// TwinCAT 3 PLC project Untitled1
// ProgramVersion: 3.1.4024.0
// libraries:
//   Tc2_Math, * (Beckhoff Automation GmbH)
//   Tc2_Standard, * (Beckhoff Automation GmbH)
//   Tc2_System, * (Beckhoff Automation GmbH)
//   Tc3_Module, * (Beckhoff Automation GmbH)
//   Tc2_MC2, * (Beckhoff Automation GmbH)
//   Tc2_MC2_Camming, * (Beckhoff Automation GmbH)
// project tree:
//   DUTs/ E_CamApplicationError.TcDUT, E_CamErrorSource.TcDUT, E_CamMachineState.TcDUT, E_CamProcessPhase.TcDUT, ST_CamCommands.TcDUT, ST_CamDerivedGeometry.TcDUT, ST_CamRecipe.TcDUT, ST_CamScope.TcDUT, ST_CamStatus.TcDUT
//   GVLs/ GVL_CamControl.TcGVL, GVL_Motion.TcGVL
//   / PlcTask.TcTTO (not stored)
//   POUs/Cam/ FB_CamMachine.TcPOU, FB_CamProfileBuilder.TcPOU, FB_CamRecipeValidator.TcPOU, FB_ElectronicCam.TcPOU, F_MakeCamPoint.TcPOU
//   POUs/Axis_test/ Axis_test.TcPOU, FB_AxisPositionTest.TcPOU
//   POUs/ MAIN.TcPOU
// real-time tasks:
//   TASK PlcTask: cycle T#10ms, priority 20, ADS port 350
// motion (NC):
//   TASK NC-Task 1 SAF: cycle T#2ms, priority 4, ADS port 501
//   TASK NC-Task 1 SVB: cycle T#10ms, priority 8, ADS port 511
//   AXIS Axis 1 (id 1)
//     OtherSettings: AllowMotionCmdToSlave=true
//     encoder EncType=19
//       EncPara: MaxCount=#xffffffff
//     drive DrvType=16
//       DrvPara: MaxCount=#xffffffff
//         Analog: TorqueSetpointScale=10, ScaleFactorActTorque=0.1
//         TimeComp: TaskDelayCycles=1
//     controller CtrType=1
//       CtrPara: PriorControlFactor=1
//         Observer: BandWidth=20
//   AXIS Axis 2 (id 2)
//     OtherSettings: AllowMotionCmdToSlave=true
//     encoder EncType=19
//       EncPara: MaxCount=#xffffffff
//     drive DrvType=16
//       DrvPara: MaxCount=#xffffffff
//         Analog: TorqueSetpointScale=10, ScaleFactorActTorque=0.1
//         TimeComp: TaskDelayCycles=1
//     controller CtrType=1
//       CtrPara: PriorControlFactor=1
//         Observer: BandWidth=20
// I/O:
//   DEVICE Device 3 (EtherCAT), AmsNetId 5.57.253.57.4.1
//     Drive 1 (INVT_DA180_114) [DA180-N EtherCAT(CoE) Drive]
//     Drive 2 (INVT_DA200A_EtherCAT_101) [INVT_DA200A_EtherCAT_1.0.1.0]
//     Term 3 (EK1100) [EK1100 EtherCAT Coupler (2A E-Bus)]
//       Term 4 (EL3164) [EL3164 4Ch. Ana. Input 0-10V]
//       Term 5 (EL9011) [EL9011 End Terminal]
// variable links:
//   NC-Task 1 SAF/Axes/Axis 1 <-> Device 3 (EtherCAT)/Drive 1 (INVT_DA180_114)
//     Drive/Inputs/In/nDataIn3[0] <-> DI Inputs/Torque Actual Value
//     Drive/Inputs/In/nDcOutputTime <-> InfoData/DcOutputShift
//     Drive/Inputs/In/nState1 <-> DI Inputs/Status Word
//     Drive/Inputs/In/nState2 <-> DI Inputs/Status Word @bit 8
//     Drive/Inputs/In/nState4 @bit 1 <-> WcState/InputToggle
//     Drive/Inputs/In/nState4 <-> WcState/WcState
//     Drive/Inputs/In/nState5 <-> DI Inputs/Operation Mode Display
//     Drive/Outputs/Out/nCtrl1 <-> DO Outputs/Control Word
//     Drive/Outputs/Out/nCtrl2 <-> DO Outputs/Control Word @bit 8
//     Drive/Outputs/Out/nCtrl5 <-> DO Outputs/Mode of Operation
//     Drive/Outputs/Out/nDataOut1 <-> DO Outputs/Target Position
//     Drive/Outputs/Out/nDataOut2 <-> DO Outputs/Target Velocity
//     Drive/Outputs/Out/nDataOut4[0] <-> DO Outputs/Target torque
//     Enc/Inputs/In/nDataIn1 <-> DI Inputs/Position Actual Value
//     Enc/Inputs/In/nDataIn3 <-> DI Inputs/Touch Probe Value
//     Enc/Inputs/In/nDataIn7 <-> DI Inputs/Speed Actual Value
//     Enc/Inputs/In/nDcInputTime <-> InfoData/DcInputShift
//     Enc/Inputs/In/nState4 @bit 1 <-> WcState/InputToggle
//     Enc/Inputs/In/nState4 <-> WcState/WcState
//     Enc/Inputs/In/nState5 <-> DI Inputs/Touch Probe Status
//     Enc/Inputs/In/nState6 <-> DI Inputs/Touch Probe Status @bit 8
//     Enc/Outputs/Out/nCtrl5 <-> DO Outputs/Touch probe control
//     Enc/Outputs/Out/nCtrl6 <-> DO Outputs/Touch probe control @bit 8
//   NC-Task 1 SAF/Axes/Axis 2 <-> Device 3 (EtherCAT)/Drive 2 (INVT_DA200A_EtherCAT_101)
//     Drive/Inputs/In/nDataIn3[0] <-> Inputs/Torque Actual Value
//     Drive/Inputs/In/nDcOutputTime <-> InfoData/DcOutputShift
//     Drive/Inputs/In/nState1 <-> Inputs/Status Word
//     Drive/Inputs/In/nState2 <-> Inputs/Status Word @bit 8
//     Drive/Inputs/In/nState4 @bit 1 <-> WcState/InputToggle
//     Drive/Inputs/In/nState4 <-> WcState/WcState
//     Drive/Inputs/In/nState5 <-> Inputs/Operation Mode Display
//     Drive/Outputs/Out/nCtrl1 <-> Outputs/Control Word
//     Drive/Outputs/Out/nCtrl2 <-> Outputs/Control Word @bit 8
//     Drive/Outputs/Out/nCtrl5 <-> Outputs/Mode of Operation
//     Drive/Outputs/Out/nDataOut1 <-> Outputs/Target Position
//     Drive/Outputs/Out/nDataOut2 <-> Outputs/Target Velocity
//     Drive/Outputs/Out/nDataOut4[0] <-> Outputs/Target torque
//     Enc/Inputs/In/nDataIn1 <-> Inputs/Position Actual Value
//     Enc/Inputs/In/nDataIn3 <-> Inputs/Touch Probe 1 Positive value
//     Enc/Inputs/In/nDataIn7 <-> Inputs/Velocity Actual Value
//     Enc/Inputs/In/nDcInputTime <-> InfoData/DcInputShift
//     Enc/Inputs/In/nState4 @bit 1 <-> WcState/InputToggle
//     Enc/Inputs/In/nState4 <-> WcState/WcState
//     Enc/Inputs/In/nState5 <-> Inputs/Touch Probe Status
//     Enc/Inputs/In/nState6 <-> Inputs/Touch Probe Status @bit 8
//     Enc/Outputs/Out/nCtrl5 <-> Outputs/Touch probe control
//     Enc/Outputs/Out/nCtrl6 <-> Outputs/Touch probe control @bit 8
//   Untitled1/Untitled1 Instance <-> NC-Task 1 SAF/Axes/Axis 1
//     PlcTask Inputs/GVL_Motion.gAxisConveyor.NcToPlc <-> Outputs/ToPlc
//     PlcTask Outputs/GVL_Motion.gAxisConveyor.PlcToNc <-> Inputs/FromPlc
//   Untitled1/Untitled1 Instance <-> NC-Task 1 SAF/Axes/Axis 2
//     PlcTask Inputs/GVL_Motion.gAxisCutter.NcToPlc <-> Outputs/ToPlc
//     PlcTask Outputs/GVL_Motion.gAxisCutter.PlcToNc <-> Inputs/FromPlc

// ---- DUTs/E_CamApplicationError.TcDUT
TYPE E_CamApplicationError :
(
    CAM_ERROR_NONE := 0,
    CAM_ERROR_COMMAND_NOT_ALLOWED,
    CAM_ERROR_NOT_REFERENCED,
    CAM_ERROR_RECIPE_PITCH,
    CAM_ERROR_RECIPE_CONVEYOR_VELOCITY,
    CAM_ERROR_RECIPE_CUT_VELOCITY,
    CAM_ERROR_RECIPE_EDGE_LENGTH,
    CAM_ERROR_RECIPE_PHASE_ORDER,
    CAM_ERROR_RECIPE_SYNC_SPACE,
    CAM_ERROR_RECIPE_RETURN_SPACE,
    CAM_ERROR_RECIPE_DYNAMICS,
    CAM_ERROR_AXIS_POWER,
    CAM_ERROR_AXIS_REFERENCE,
    CAM_ERROR_CAM_BUILD,
    CAM_ERROR_CAM_LOAD,
    CAM_ERROR_CAM_CHARACTERISTICS,
    CAM_ERROR_CAM_IN,
    CAM_ERROR_MASTER_MOVE,
    CAM_ERROR_MASTER_STOP,
    CAM_ERROR_CAM_OUT,
    CAM_ERROR_SLAVE_RETURN,
    CAM_ERROR_AXIS_RESET
);
END_TYPE

// ---- DUTs/E_CamErrorSource.TcDUT
TYPE E_CamErrorSource :
(
    CAM_SOURCE_NONE := 0,
    CAM_SOURCE_RECIPE,
    CAM_SOURCE_MASTER_AXIS,
    CAM_SOURCE_SLAVE_AXIS,
    CAM_SOURCE_TABLE_LOAD,
    CAM_SOURCE_TABLE_CHARACTERISTICS,
    CAM_SOURCE_CAM_IN,
    CAM_SOURCE_CAM_OUT
);
END_TYPE

// ---- DUTs/E_CamMachineState.TcDUT
TYPE E_CamMachineState :
(
    CAM_STATE_DISABLED := 0,
    CAM_STATE_POWERING,
    CAM_STATE_IDLE,
    CAM_STATE_REFERENCING_MASTER,
    CAM_STATE_REFERENCING_SLAVE,
    CAM_STATE_BUILDING_TABLE,
    CAM_STATE_LOADING_TABLE,
    CAM_STATE_READY,
    CAM_STATE_CAMMING_IN,
    CAM_STATE_STARTING_MASTER,
    CAM_STATE_RUNNING,
    CAM_STATE_STOPPING_MASTER,
    CAM_STATE_RELEASING_STOP,
    CAM_STATE_CAMMING_OUT,
    CAM_STATE_RETURNING_SLAVE,
    CAM_STATE_RESETTING,
    CAM_STATE_FAULT
);
END_TYPE

// ---- DUTs/E_CamProcessPhase.TcDUT
TYPE E_CamProcessPhase :
(
    CAM_PHASE_DISABLED := 0,
    CAM_PHASE_PREPARE,
    CAM_PHASE_APPROACH,
    CAM_PHASE_FIRST_EDGE,
    CAM_PHASE_EXIT_FIRST_EDGE,
    CAM_PHASE_SYNCHRONOUS,
    CAM_PHASE_ENTER_SECOND_EDGE,
    CAM_PHASE_SECOND_EDGE,
    CAM_PHASE_RETURN,
    CAM_PHASE_DWELL
);
END_TYPE

// ---- DUTs/ST_CamCommands.TcDUT
TYPE ST_CamCommands :
STRUCT
    bEnable : BOOL;
    bReference : BOOL;
    bApplyRecipe : BOOL;
    bStart : BOOL;
    bStop : BOOL;
    bReset : BOOL;
END_STRUCT
END_TYPE

// ---- DUTs/ST_CamDerivedGeometry.TcDUT
TYPE ST_CamDerivedGeometry :
STRUCT
    lrCutMasterDistance : LREAL;
    lrFirstSlope : LREAL;
    lrSecondSlope : LREAL;
    lrFirstEdgeEnd : LREAL;
    lrExitBlendEnd : LREAL;
    lrEntryBlendStart : LREAL;
    lrSecondEdgeEnd : LREAL;
    lrClearanceRelative : LREAL;
    lrFirstStartY : LREAL;
    lrFirstEndY : LREAL;
    lrExitEndY : LREAL;
    lrEntryStartY : LREAL;
    lrSecondStartY : LREAL;
    lrSecondEndY : LREAL;
    lrMasterStopDistance : LREAL;
    lrStopWindowMargin : LREAL;
END_STRUCT
END_TYPE

// ---- DUTs/ST_CamRecipe.TcDUT
TYPE ST_CamRecipe :
STRUCT
    lrObjectPitch : LREAL := 500.0;
    lrConveyorVelocity : LREAL := 100.0;
    lrCutVelocity : LREAL := 50.0;
    lrObjectEdgeLength : LREAL := 25.0;
    lrFirstEdgeStart : LREAL := 100.0;
    lrSecondEdgeStart : LREAL := 300.0;
    lrBlendMasterDistance : LREAL := 20.0;
    lrReturnEndPhase : LREAL := 480.0;
    lrMasterAcceleration : LREAL := 500.0;
    lrMasterDeceleration : LREAL := 500.0;
    lrMasterJerk : LREAL := 5000.0;
    lrMaxSlaveVelocity : LREAL := 600.0;
    lrMaxSlaveAcceleration : LREAL := 1600.0;
    lrMaxSlaveJerk : LREAL := 12000.0;
    lrRecoveryVelocity : LREAL := 100.0;
    lrRecoveryAcceleration : LREAL := 500.0;
    lrRecoveryDeceleration : LREAL := 500.0;
    lrRecoveryJerk : LREAL := 5000.0;
    lrPositionTolerance : LREAL := 0.1;
END_STRUCT
END_TYPE

// ---- DUTs/ST_CamScope.TcDUT
TYPE ST_CamScope :
STRUCT
    lrMasterSetPosition : LREAL;
    lrMasterActualPosition : LREAL;
    lrMasterSetVelocity : LREAL;
    lrMasterActualVelocity : LREAL;
    lrMasterPhase : LREAL;
    lrSlaveSetPosition : LREAL;
    lrSlaveActualPosition : LREAL;
    lrSlaveSetVelocity : LREAL;
    lrSlaveActualVelocity : LREAL;
    lrExpectedSlaveVelocity : LREAL;
    lrObjectRelativePosition : LREAL;
    eMachineState : E_CamMachineState;
    eProcessPhase : E_CamProcessPhase;
    bCamActive : BOOL;
    bRecipeLoaded : BOOL;
    eApplicationError : E_CamApplicationError;
    udiMotionErrorID : UDINT;
END_STRUCT
END_TYPE

// ---- DUTs/ST_CamStatus.TcDUT
TYPE ST_CamStatus :
STRUCT
    eState : E_CamMachineState;
    eProcessPhase : E_CamProcessPhase;
    bPowerEnabled : BOOL;
    bReferenced : BOOL;
    bRecipeLoaded : BOOL;
    bCamActive : BOOL;
    bRunning : BOOL;
    bBusy : BOOL;
    eApplicationError : E_CamApplicationError;
    eErrorSource : E_CamErrorSource;
    udiMotionErrorID : UDINT;
    lrCalculatedMaxSlaveVelocity : LREAL;
    lrCalculatedMaxSlaveAcceleration : LREAL;
    lrCalculatedMaxSlaveJerk : LREAL;
    lrCalculatedFaultStopSlaveAcceleration : LREAL;
    lrCalculatedFaultStopSlaveJerk : LREAL;
END_STRUCT
END_TYPE

// ---- GVLs/GVL_CamControl.TcGVL
{attribute 'qualified_only'}
VAR_GLOBAL
    stCommands : ST_CamCommands;
    stRecipe : ST_CamRecipe;
    stStatus : ST_CamStatus;
    stScope : ST_CamScope;
END_VAR

// ---- GVLs/GVL_Motion.TcGVL
{attribute 'qualified_only'}
VAR_GLOBAL
    gAxisConveyor : AXIS_REF;
    gAxisCutter : AXIS_REF;
END_VAR

// ---- POUs/Cam/FB_CamMachine.TcPOU
FUNCTION_BLOCK FB_CamMachine
VAR_INPUT
    stCommands : ST_CamCommands;
    stRecipe : ST_CamRecipe;
END_VAR
VAR_IN_OUT
    AxisConveyor : AXIS_REF;
    AxisCutter : AXIS_REF;
END_VAR
VAR_OUTPUT
    stStatus : ST_CamStatus;
    stScope : ST_CamScope;
END_VAR
VAR CONSTANT
    c_nCamTableIdA : MC_CAM_ID := 1;
    c_nCamTableIdB : MC_CAM_ID := 2;
    // Commissioned application limits; NC/drive limits must be no lower.
    c_lrMachineMaxSlaveVelocity : LREAL := 600.0;
    c_lrMachineMaxSlaveAcceleration : LREAL := 1600.0;
    c_lrMachineMaxSlaveJerk : LREAL := 12000.0;
    // Conservative controlled stop used only after a runtime fault.
    c_lrFaultStopDeceleration : LREAL := 15.0;
    c_lrFaultStopJerk : LREAL := 50.0;
END_VAR
VAR
    eState : E_CamMachineState := CAM_STATE_DISABLED;
    eProcessPhase : E_CamProcessPhase := CAM_PHASE_DISABLED;

    rtReference : R_TRIG;
    rtApplyRecipe : R_TRIG;
    rtStart : R_TRIG;
    rtStop : R_TRIG;
    rtReset : R_TRIG;

    fbPowerConveyor : MC_Power;
    fbPowerCutter : MC_Power;
    fbSetPositionConveyor : MC_SetPosition;
    fbSetPositionCutter : MC_SetPosition;
    fbResetConveyor : MC_Reset;
    fbResetCutter : MC_Reset;
    fbMoveConveyor : MC_MoveVelocity;
    fbStopConveyor : MC_Stop;
    fbReturnCutter : MC_MoveAbsolute;

    fbRecipeValidator : FB_CamRecipeValidator;
    fbProfileBuilder : FB_CamProfileBuilder;
    fbElectronicCam : FB_ElectronicCam;

    stPowerOptions : ST_PowerOptions;
    stSetPositionConveyorOptions : ST_SetPositionOptions;
    stSetPositionCutterOptions : ST_SetPositionOptions;
    stMoveConveyorOptions : ST_MoveOptions;
    stStopConveyorOptions : ST_MoveOptions;
    stReturnCutterOptions : ST_MoveOptions;

    stPendingRecipe : ST_CamRecipe;
    stActiveRecipe : ST_CamRecipe;
    stDerived : ST_CamDerivedGeometry;
    stCamRef : MC_CAM_REF;

    bPowerRequest : BOOL;
    bReferenced : BOOL;
    bRecipeLoaded : BOOL;
    bStopRequested : BOOL;
    bResetInProgress : BOOL;
    bFaultStop : BOOL;
    bForcePowerOff : BOOL;
    usiBuildState : USINT;

    nActiveCamTableId : MC_CAM_ID := 1;
    nCandidateCamTableId : MC_CAM_ID := 2;
    nCamCommandTableId : MC_CAM_ID := 1;

    bSetPositionConveyorExecute : BOOL;
    bSetPositionCutterExecute : BOOL;
    bResetConveyorExecute : BOOL;
    bResetCutterExecute : BOOL;
    bMoveConveyorExecute : BOOL;
    bStopConveyorExecute : BOOL;
    bReturnCutterExecute : BOOL;

    bValidateRecipePulse : BOOL;
    bBuildProfilePulse : BOOL;
    bLoadCamPulse : BOOL;
    bCoupleCamPulse : BOOL;
    bDecoupleCamPulse : BOOL;
    bResetCamPulse : BOOL;

    lrMasterCycleOrigin : LREAL;
    lrMasterPhase : LREAL;
    lrSlaveCycleOrigin : LREAL;
    lrSlaveCamPosition : LREAL;
    lrStopCommandDeceleration : LREAL;
    lrStopCommandJerk : LREAL;
    lrMaxCamSlope : LREAL;
    lrMaxCamSecondDerivative : LREAL;
    lrCalculatedMaxSlaveVelocity : LREAL;
    lrCalculatedMaxSlaveAcceleration : LREAL;
    lrCalculatedMaxSlaveJerk : LREAL;
    lrCalculatedFaultStopSlaveAcceleration : LREAL;
    lrCalculatedFaultStopSlaveJerk : LREAL;

    bFaultLatched : BOOL;
    eLatchedApplicationError : E_CamApplicationError;
    eLatchedErrorSource : E_CamErrorSource;
    udiLatchedMotionErrorID : UDINT;
    bRequestFault : BOOL;
    eRequestedApplicationError : E_CamApplicationError;
    eRequestedErrorSource : E_CamErrorSource;
    udiRequestedMotionErrorID : UDINT;
END_VAR

// Refresh both axis status structures once at the start of the PLC scan.
AxisConveyor.ReadStatus();
AxisCutter.ReadStatus();

rtReference(CLK := stCommands.bReference);
rtApplyRecipe(CLK := stCommands.bApplyRecipe);
rtStart(CLK := stCommands.bStart);
rtStop(CLK := stCommands.bStop);
rtReset(CLK := stCommands.bReset);

// One-scan requests consumed by the lower layers at the end of this call.
bValidateRecipePulse := FALSE;
bBuildProfilePulse := FALSE;
bLoadCamPulse := FALSE;
bCoupleCamPulse := FALSE;
bDecoupleCamPulse := FALSE;
bResetCamPulse := FALSE;

bRequestFault := FALSE;
eRequestedApplicationError := CAM_ERROR_NONE;
eRequestedErrorSource := CAM_SOURCE_NONE;
udiRequestedMotionErrorID := 0;

IF stActiveRecipe.lrObjectPitch > 0.0 THEN
    lrMasterPhase := MODABS(
        AxisConveyor.NcToPlc.SetPos - lrMasterCycleOrigin,
        stActiveRecipe.lrObjectPitch);
ELSE
    lrMasterPhase := 0.0;
END_IF;

CASE eState OF
    CAM_STATE_DISABLED:
        bSetPositionConveyorExecute := FALSE;
        bSetPositionCutterExecute := FALSE;
        bResetConveyorExecute := FALSE;
        bResetCutterExecute := FALSE;
        bMoveConveyorExecute := FALSE;
        bStopConveyorExecute := FALSE;
        bReturnCutterExecute := FALSE;
        bStopRequested := FALSE;
        IF stCommands.bEnable THEN
            eState := CAM_STATE_POWERING;
        END_IF;

    CAM_STATE_POWERING:
        IF NOT stCommands.bEnable THEN
            eState := CAM_STATE_DISABLED;
        ELSIF fbPowerConveyor.Status AND fbPowerCutter.Status THEN
            IF bReferenced AND bRecipeLoaded THEN
                eState := CAM_STATE_READY;
            ELSE
                eState := CAM_STATE_IDLE;
            END_IF;
        END_IF;

    CAM_STATE_IDLE:
        IF NOT stCommands.bEnable THEN
            eState := CAM_STATE_DISABLED;
        ELSIF rtReference.Q THEN
            IF AxisConveyor.Status.NotMoving AND AxisCutter.Status.NotMoving THEN
                bReferenced := FALSE;
                bRecipeLoaded := FALSE;
                bSetPositionConveyorExecute := TRUE;
                eState := CAM_STATE_REFERENCING_MASTER;
            ELSE
                bRequestFault := TRUE;
                eRequestedApplicationError := CAM_ERROR_COMMAND_NOT_ALLOWED;
            END_IF;
        ELSIF rtApplyRecipe.Q THEN
            IF NOT bReferenced THEN
                bRequestFault := TRUE;
                eRequestedApplicationError := CAM_ERROR_NOT_REFERENCED;
                eRequestedErrorSource := CAM_SOURCE_RECIPE;
            ELSIF AxisConveyor.Status.NotMoving
               AND AxisCutter.Status.NotMoving
               AND NOT fbElectronicCam.bCamActive THEN
                stPendingRecipe := stRecipe;
                IF nActiveCamTableId = c_nCamTableIdA THEN
                    nCandidateCamTableId := c_nCamTableIdB;
                ELSE
                    nCandidateCamTableId := c_nCamTableIdA;
                END_IF;
                nCamCommandTableId := nCandidateCamTableId;
                bRecipeLoaded := FALSE;
                usiBuildState := 0;
                eState := CAM_STATE_BUILDING_TABLE;
            ELSE
                bRequestFault := TRUE;
                eRequestedApplicationError := CAM_ERROR_COMMAND_NOT_ALLOWED;
            END_IF;
        ELSIF rtStart.Q THEN
            bRequestFault := TRUE;
            eRequestedApplicationError := CAM_ERROR_COMMAND_NOT_ALLOWED;
        END_IF;

    CAM_STATE_REFERENCING_MASTER:
        IF fbSetPositionConveyor.Done THEN
            bSetPositionConveyorExecute := FALSE;
            bSetPositionCutterExecute := TRUE;
            eState := CAM_STATE_REFERENCING_SLAVE;
        END_IF;

    CAM_STATE_REFERENCING_SLAVE:
        IF fbSetPositionCutter.Done THEN
            bSetPositionCutterExecute := FALSE;
            bReferenced := TRUE;
            eState := CAM_STATE_IDLE;
        END_IF;

    CAM_STATE_BUILDING_TABLE:
        IF rtReference.Q OR rtApplyRecipe.Q OR rtStart.Q THEN
            bRequestFault := TRUE;
            eRequestedApplicationError := CAM_ERROR_COMMAND_NOT_ALLOWED;
        END_IF;

        CASE usiBuildState OF
            0:
                bValidateRecipePulse := TRUE;
                usiBuildState := 10;

            10:
                IF fbRecipeValidator.bDone THEN
                    IF fbRecipeValidator.bValid THEN
                        stDerived := fbRecipeValidator.stDerived;
                        bBuildProfilePulse := TRUE;
                        usiBuildState := 20;
                    ELSE
                        bRequestFault := TRUE;
                        eRequestedApplicationError := fbRecipeValidator.eError;
                        eRequestedErrorSource := CAM_SOURCE_RECIPE;
                    END_IF;
                END_IF;

            20:
                IF fbProfileBuilder.bDone THEN
                    stCamRef := fbProfileBuilder.stCamRef;
                    bLoadCamPulse := TRUE;
                    usiBuildState := 0;
                    eState := CAM_STATE_LOADING_TABLE;
                END_IF;
        END_CASE;

    CAM_STATE_LOADING_TABLE:
        IF rtReference.Q OR rtApplyRecipe.Q OR rtStart.Q THEN
            bRequestFault := TRUE;
            eRequestedApplicationError := CAM_ERROR_COMMAND_NOT_ALLOWED;
        ELSIF fbElectronicCam.bLoadDone THEN
            lrCalculatedMaxSlaveVelocity := MAX(
                ABS(fbElectronicCam.stCharacteristics.fSlaveVeloMin),
                ABS(fbElectronicCam.stCharacteristics.fSlaveVeloMax))
                * stPendingRecipe.lrConveyorVelocity;
            lrCalculatedMaxSlaveAcceleration := MAX(
                ABS(fbElectronicCam.stCharacteristics.fSlaveAccMin),
                ABS(fbElectronicCam.stCharacteristics.fSlaveAccMax))
                * stPendingRecipe.lrConveyorVelocity
                * stPendingRecipe.lrConveyorVelocity;
            lrCalculatedMaxSlaveJerk := MAX(
                ABS(fbElectronicCam.stCharacteristics.fSlaveJerkMin),
                ABS(fbElectronicCam.stCharacteristics.fSlaveJerkMax))
                * stPendingRecipe.lrConveyorVelocity
                * stPendingRecipe.lrConveyorVelocity
                * stPendingRecipe.lrConveyorVelocity;
            lrMaxCamSlope := MAX(
                ABS(fbElectronicCam.stCharacteristics.fSlaveVeloMin),
                ABS(fbElectronicCam.stCharacteristics.fSlaveVeloMax));
            lrMaxCamSecondDerivative := MAX(
                ABS(fbElectronicCam.stCharacteristics.fSlaveAccMin),
                ABS(fbElectronicCam.stCharacteristics.fSlaveAccMax));
            lrCalculatedFaultStopSlaveAcceleration :=
                lrCalculatedMaxSlaveAcceleration
                + lrMaxCamSlope * c_lrFaultStopDeceleration;
            lrCalculatedFaultStopSlaveJerk :=
                lrCalculatedMaxSlaveJerk
                + 3.0 * lrMaxCamSecondDerivative
                  * stPendingRecipe.lrConveyorVelocity
                  * c_lrFaultStopDeceleration
                + lrMaxCamSlope * c_lrFaultStopJerk;

            IF (lrCalculatedMaxSlaveVelocity > stPendingRecipe.lrMaxSlaveVelocity)
               OR (lrCalculatedMaxSlaveAcceleration
                    > stPendingRecipe.lrMaxSlaveAcceleration)
               OR (lrCalculatedMaxSlaveJerk > stPendingRecipe.lrMaxSlaveJerk)
               OR (lrCalculatedFaultStopSlaveAcceleration
                    > stPendingRecipe.lrMaxSlaveAcceleration)
               OR (lrCalculatedFaultStopSlaveJerk
                    > stPendingRecipe.lrMaxSlaveJerk)
               OR (lrCalculatedMaxSlaveVelocity
                    > c_lrMachineMaxSlaveVelocity)
               OR (lrCalculatedMaxSlaveAcceleration
                    > c_lrMachineMaxSlaveAcceleration)
               OR (lrCalculatedMaxSlaveJerk > c_lrMachineMaxSlaveJerk)
               OR (lrCalculatedFaultStopSlaveAcceleration
                    > c_lrMachineMaxSlaveAcceleration)
               OR (lrCalculatedFaultStopSlaveJerk
                    > c_lrMachineMaxSlaveJerk) THEN
                bRequestFault := TRUE;
                eRequestedApplicationError := CAM_ERROR_RECIPE_DYNAMICS;
                eRequestedErrorSource := CAM_SOURCE_TABLE_CHARACTERISTICS;
            ELSE
                stActiveRecipe := stPendingRecipe;
                nActiveCamTableId := nCandidateCamTableId;
                nCamCommandTableId := nActiveCamTableId;
                bRecipeLoaded := TRUE;
                IF stCommands.bEnable THEN
                    eState := CAM_STATE_READY;
                ELSE
                    eState := CAM_STATE_DISABLED;
                END_IF;
            END_IF;
        END_IF;

    CAM_STATE_READY:
        bStopRequested := FALSE;
        bFaultStop := FALSE;
        IF NOT stCommands.bEnable THEN
            eState := CAM_STATE_DISABLED;
        ELSIF rtReference.Q THEN
            IF AxisConveyor.Status.NotMoving AND AxisCutter.Status.NotMoving THEN
                bReferenced := FALSE;
                bRecipeLoaded := FALSE;
                bSetPositionConveyorExecute := TRUE;
                eState := CAM_STATE_REFERENCING_MASTER;
            ELSE
                bRequestFault := TRUE;
                eRequestedApplicationError := CAM_ERROR_COMMAND_NOT_ALLOWED;
            END_IF;
        ELSIF rtApplyRecipe.Q THEN
            IF NOT bReferenced THEN
                bRequestFault := TRUE;
                eRequestedApplicationError := CAM_ERROR_NOT_REFERENCED;
                eRequestedErrorSource := CAM_SOURCE_RECIPE;
            ELSIF AxisConveyor.Status.NotMoving
               AND AxisCutter.Status.NotMoving
               AND NOT fbElectronicCam.bCamActive THEN
                stPendingRecipe := stRecipe;
                IF nActiveCamTableId = c_nCamTableIdA THEN
                    nCandidateCamTableId := c_nCamTableIdB;
                ELSE
                    nCandidateCamTableId := c_nCamTableIdA;
                END_IF;
                nCamCommandTableId := nCandidateCamTableId;
                bRecipeLoaded := FALSE;
                usiBuildState := 0;
                eState := CAM_STATE_BUILDING_TABLE;
            ELSE
                bRequestFault := TRUE;
                eRequestedApplicationError := CAM_ERROR_COMMAND_NOT_ALLOWED;
            END_IF;
        ELSIF rtStart.Q THEN
            IF bReferenced
               AND bRecipeLoaded
               AND AxisConveyor.Status.NotMoving
               AND AxisCutter.Status.NotMoving
               AND NOT fbElectronicCam.bCamActive
               AND (ABS(AxisCutter.NcToPlc.SetPos)
                    <= stActiveRecipe.lrPositionTolerance) THEN
                bStopRequested := FALSE;
                bFaultStop := FALSE;
                bMoveConveyorExecute := TRUE;
                eState := CAM_STATE_STARTING_MASTER;
            ELSE
                bRequestFault := TRUE;
                eRequestedApplicationError := CAM_ERROR_COMMAND_NOT_ALLOWED;
            END_IF;
        END_IF;

    CAM_STATE_STARTING_MASTER:
        IF rtStop.Q OR NOT stCommands.bEnable THEN
            bMoveConveyorExecute := FALSE;
            bFaultStop := FALSE;
            bStopConveyorExecute := TRUE;
            eState := CAM_STATE_STOPPING_MASTER;
        ELSIF rtReference.Q OR rtApplyRecipe.Q OR rtStart.Q THEN
            bRequestFault := TRUE;
            eRequestedApplicationError := CAM_ERROR_COMMAND_NOT_ALLOWED;
        ELSIF fbMoveConveyor.InVelocity THEN
            // Cam coupling starts only after the conveyor is at constant speed.
            bMoveConveyorExecute := FALSE;
            lrMasterCycleOrigin := AxisConveyor.NcToPlc.SetPos;
            lrSlaveCycleOrigin := AxisCutter.NcToPlc.SetPos;
            nCamCommandTableId := nActiveCamTableId;
            bCoupleCamPulse := TRUE;
            eState := CAM_STATE_CAMMING_IN;
        END_IF;

    CAM_STATE_CAMMING_IN:
        IF rtStop.Q OR NOT stCommands.bEnable THEN
            bStopRequested := TRUE;
        END_IF;
        IF rtReference.Q OR rtApplyRecipe.Q OR rtStart.Q THEN
            bStopRequested := TRUE;
            bRequestFault := TRUE;
            eRequestedApplicationError := CAM_ERROR_COMMAND_NOT_ALLOWED;
        END_IF;
        IF fbElectronicCam.bError THEN
            IF NOT bFaultLatched THEN
                bRequestFault := TRUE;
                eRequestedApplicationError := fbElectronicCam.eApplicationError;
                eRequestedErrorSource := fbElectronicCam.eErrorSource;
                udiRequestedMotionErrorID := fbElectronicCam.udiErrorID;
            END_IF;
        ELSIF fbElectronicCam.bCoupleDone THEN
            IF bStopRequested OR bFaultLatched OR bRequestFault THEN
                bFaultStop := bFaultLatched OR bRequestFault;
                eState := CAM_STATE_STOPPING_MASTER;
            ELSE
                eState := CAM_STATE_RUNNING;
            END_IF;
        END_IF;

    CAM_STATE_RUNNING:
        IF rtStop.Q OR NOT stCommands.bEnable THEN
            bStopRequested := TRUE;
            bFaultStop := FALSE;
            eState := CAM_STATE_STOPPING_MASTER;
        ELSIF rtReference.Q OR rtApplyRecipe.Q OR rtStart.Q THEN
            bRequestFault := TRUE;
            eRequestedApplicationError := CAM_ERROR_COMMAND_NOT_ALLOWED;
        END_IF;

    CAM_STATE_STOPPING_MASTER:
        IF rtReference.Q OR rtApplyRecipe.Q OR rtStart.Q THEN
            bRequestFault := TRUE;
            eRequestedApplicationError := CAM_ERROR_COMMAND_NOT_ALLOWED;
        END_IF;

        // A normal stop waits for the zero-slope 480..500 mm dwell. A fault
        // stop uses the separately validated conservative dynamics immediately.
        IF NOT bStopConveyorExecute THEN
            IF bFaultStop OR NOT fbElectronicCam.bCamActive THEN
                bStopConveyorExecute := TRUE;
            ELSIF (lrMasterPhase >= stActiveRecipe.lrReturnEndPhase)
               AND (lrMasterPhase <=
                    (stActiveRecipe.lrObjectPitch
                     - stDerived.lrMasterStopDistance
                     - stDerived.lrStopWindowMargin)) THEN
                bStopConveyorExecute := TRUE;
            END_IF;
        END_IF;

        IF fbStopConveyor.Error THEN
            bStopConveyorExecute := FALSE;
            bRequestFault := TRUE;
            eRequestedApplicationError := CAM_ERROR_MASTER_STOP;
            eRequestedErrorSource := CAM_SOURCE_MASTER_AXIS;
            udiRequestedMotionErrorID := fbStopConveyor.ErrorID;
            bForcePowerOff := TRUE;
            eState := CAM_STATE_FAULT;
        ELSIF fbStopConveyor.Done THEN
            bStopConveyorExecute := FALSE;
            eState := CAM_STATE_RELEASING_STOP;
        END_IF;

    CAM_STATE_RELEASING_STOP:
        IF rtReference.Q OR rtApplyRecipe.Q OR rtStart.Q THEN
            bRequestFault := TRUE;
            eRequestedApplicationError := CAM_ERROR_COMMAND_NOT_ALLOWED;
        END_IF;
        IF NOT fbStopConveyor.Busy THEN
            IF fbElectronicCam.bCamActive THEN
                bDecoupleCamPulse := TRUE;
                eState := CAM_STATE_CAMMING_OUT;
            ELSE
                bReturnCutterExecute := TRUE;
                eState := CAM_STATE_RETURNING_SLAVE;
            END_IF;
        END_IF;

    CAM_STATE_CAMMING_OUT:
        IF rtReference.Q OR rtApplyRecipe.Q OR rtStart.Q THEN
            bRequestFault := TRUE;
            eRequestedApplicationError := CAM_ERROR_COMMAND_NOT_ALLOWED;
        END_IF;
        IF fbElectronicCam.bError THEN
            IF NOT bFaultLatched THEN
                bRequestFault := TRUE;
                eRequestedApplicationError := fbElectronicCam.eApplicationError;
                eRequestedErrorSource := fbElectronicCam.eErrorSource;
                udiRequestedMotionErrorID := fbElectronicCam.udiErrorID;
            END_IF;
            eState := CAM_STATE_FAULT;
        ELSIF fbElectronicCam.bDecoupleDone THEN
            bReturnCutterExecute := TRUE;
            eState := CAM_STATE_RETURNING_SLAVE;
        END_IF;

    CAM_STATE_RETURNING_SLAVE:
        IF NOT bResetInProgress
           AND (rtReference.Q OR rtApplyRecipe.Q OR rtStart.Q) THEN
            bRequestFault := TRUE;
            eRequestedApplicationError := CAM_ERROR_COMMAND_NOT_ALLOWED;
        END_IF;
        IF fbReturnCutter.Error OR fbReturnCutter.CommandAborted THEN
            bReturnCutterExecute := FALSE;
            IF NOT bFaultLatched THEN
                bRequestFault := TRUE;
                eRequestedApplicationError := CAM_ERROR_SLAVE_RETURN;
                eRequestedErrorSource := CAM_SOURCE_SLAVE_AXIS;
                udiRequestedMotionErrorID := fbReturnCutter.ErrorID;
            END_IF;
            eState := CAM_STATE_FAULT;
        ELSIF fbReturnCutter.Done
           AND (ABS(AxisCutter.NcToPlc.SetPos)
                <= stActiveRecipe.lrPositionTolerance) THEN
            bReturnCutterExecute := FALSE;
            bStopRequested := FALSE;
            IF bResetInProgress THEN
                bResetInProgress := FALSE;
                bFaultStop := FALSE;
                bForcePowerOff := FALSE;
                bFaultLatched := FALSE;
                eLatchedApplicationError := CAM_ERROR_NONE;
                eLatchedErrorSource := CAM_SOURCE_NONE;
                udiLatchedMotionErrorID := 0;
                bRecipeLoaded := FALSE;
                IF stCommands.bEnable THEN
                    eState := CAM_STATE_POWERING;
                ELSE
                    eState := CAM_STATE_DISABLED;
                END_IF;
            ELSIF bFaultLatched THEN
                eState := CAM_STATE_FAULT;
            ELSIF stCommands.bEnable THEN
                eState := CAM_STATE_READY;
            ELSE
                eState := CAM_STATE_DISABLED;
            END_IF;
        END_IF;

    CAM_STATE_RESETTING:
        IF fbResetConveyor.Error OR fbResetCutter.Error THEN
            bResetConveyorExecute := FALSE;
            bResetCutterExecute := FALSE;
            bResetInProgress := FALSE;
            eState := CAM_STATE_FAULT;
        ELSIF fbResetConveyor.Done AND fbResetCutter.Done THEN
            bResetConveyorExecute := FALSE;
            bResetCutterExecute := FALSE;
            IF fbElectronicCam.bCamActive THEN
                bDecoupleCamPulse := TRUE;
                eState := CAM_STATE_CAMMING_OUT;
            ELSE
                bReturnCutterExecute := TRUE;
                eState := CAM_STATE_RETURNING_SLAVE;
            END_IF;
        END_IF;

    CAM_STATE_FAULT:
        bSetPositionConveyorExecute := FALSE;
        bSetPositionCutterExecute := FALSE;
        bMoveConveyorExecute := FALSE;
        bStopConveyorExecute := FALSE;
        bReturnCutterExecute := FALSE;
        IF rtReset.Q
           AND AxisConveyor.Status.NotMoving
           AND AxisCutter.Status.NotMoving THEN
            bFaultStop := FALSE;
            bForcePowerOff := FALSE;
            bResetConveyorExecute := TRUE;
            bResetCutterExecute := TRUE;
            bResetCamPulse := TRUE;
            bResetInProgress := TRUE;
            eState := CAM_STATE_RESETTING;
        END_IF;
END_CASE;

// Keep power while any controlled stop, decouple, return, or reset is active.
// MC_Stop failure removes the non-safety motion enable as a last fallback.
bPowerRequest := (stCommands.bEnable
    OR (eState = CAM_STATE_REFERENCING_MASTER)
    OR (eState = CAM_STATE_REFERENCING_SLAVE)
    OR (eState = CAM_STATE_CAMMING_IN)
    OR (eState = CAM_STATE_STARTING_MASTER)
    OR (eState = CAM_STATE_RUNNING)
    OR (eState = CAM_STATE_STOPPING_MASTER)
    OR (eState = CAM_STATE_RELEASING_STOP)
    OR (eState = CAM_STATE_CAMMING_OUT)
    OR (eState = CAM_STATE_RETURNING_SLAVE)
    OR (eState = CAM_STATE_RESETTING)
    OR fbElectronicCam.bBusy
    OR fbElectronicCam.bCamActive)
    AND NOT bForcePowerOff;

fbPowerConveyor(
    Enable := bPowerRequest,
    Enable_Positive := TRUE,
    Enable_Negative := TRUE,
    Override := 100.0,
    BufferMode := MC_Aborting,
    Options := stPowerOptions,
    Axis := AxisConveyor);
fbPowerCutter(
    Enable := bPowerRequest,
    Enable_Positive := TRUE,
    Enable_Negative := TRUE,
    Override := 100.0,
    BufferMode := MC_Aborting,
    Options := stPowerOptions,
    Axis := AxisCutter);

fbSetPositionConveyor(
    Execute := bSetPositionConveyorExecute,
    Position := 0.0,
    Mode := FALSE,
    Options := stSetPositionConveyorOptions,
    Axis := AxisConveyor);
fbSetPositionCutter(
    Execute := bSetPositionCutterExecute,
    Position := 0.0,
    Mode := FALSE,
    Options := stSetPositionCutterOptions,
    Axis := AxisCutter);

fbResetConveyor(
    Execute := bResetConveyorExecute,
    Axis := AxisConveyor);
fbResetCutter(
    Execute := bResetCutterExecute,
    Axis := AxisCutter);

fbMoveConveyor(
    Execute := bMoveConveyorExecute,
    Velocity := stActiveRecipe.lrConveyorVelocity,
    Acceleration := stActiveRecipe.lrMasterAcceleration,
    Deceleration := stActiveRecipe.lrMasterDeceleration,
    Jerk := stActiveRecipe.lrMasterJerk,
    Direction := MC_Positive_Direction,
    BufferMode := MC_Aborting,
    Options := stMoveConveyorOptions,
    Axis := AxisConveyor);
IF bFaultStop THEN
    lrStopCommandDeceleration := c_lrFaultStopDeceleration;
    lrStopCommandJerk := c_lrFaultStopJerk;
ELSE
    lrStopCommandDeceleration := stActiveRecipe.lrMasterDeceleration;
    lrStopCommandJerk := stActiveRecipe.lrMasterJerk;
END_IF;
fbStopConveyor(
    Execute := bStopConveyorExecute,
    Deceleration := lrStopCommandDeceleration,
    Jerk := lrStopCommandJerk,
    Options := stStopConveyorOptions,
    Axis := AxisConveyor);
fbReturnCutter(
    Execute := bReturnCutterExecute,
    Position := 0.0,
    Velocity := stActiveRecipe.lrRecoveryVelocity,
    Acceleration := stActiveRecipe.lrRecoveryAcceleration,
    Deceleration := stActiveRecipe.lrRecoveryDeceleration,
    Jerk := stActiveRecipe.lrRecoveryJerk,
    BufferMode := MC_Aborting,
    Options := stReturnCutterOptions,
    Axis := AxisCutter);

fbRecipeValidator(
    bExecute := bValidateRecipePulse,
    stRecipe := stPendingRecipe);
fbProfileBuilder(
    bExecute := bBuildProfilePulse,
    stRecipe := stPendingRecipe,
    stDerived := stDerived);
fbElectronicCam(
    bLoad := bLoadCamPulse,
    bCouple := bCoupleCamPulse,
    bDecouple := bDecoupleCamPulse,
    bReset := bResetCamPulse,
    nCamTableId := nCamCommandTableId,
    Master := AxisConveyor,
    Slave := AxisCutter,
    CamTable := stCamRef);

// Convert lower-level errors into one deterministic first-fault request.
IF NOT bRequestFault AND NOT bFaultLatched THEN
    IF fbPowerConveyor.Error THEN
        bRequestFault := TRUE;
        eRequestedApplicationError := CAM_ERROR_AXIS_POWER;
        eRequestedErrorSource := CAM_SOURCE_MASTER_AXIS;
        udiRequestedMotionErrorID := fbPowerConveyor.ErrorID;
    ELSIF fbPowerCutter.Error THEN
        bRequestFault := TRUE;
        eRequestedApplicationError := CAM_ERROR_AXIS_POWER;
        eRequestedErrorSource := CAM_SOURCE_SLAVE_AXIS;
        udiRequestedMotionErrorID := fbPowerCutter.ErrorID;
    ELSIF fbSetPositionConveyor.Error THEN
        bRequestFault := TRUE;
        eRequestedApplicationError := CAM_ERROR_AXIS_REFERENCE;
        eRequestedErrorSource := CAM_SOURCE_MASTER_AXIS;
        udiRequestedMotionErrorID := fbSetPositionConveyor.ErrorID;
    ELSIF fbSetPositionCutter.Error THEN
        bRequestFault := TRUE;
        eRequestedApplicationError := CAM_ERROR_AXIS_REFERENCE;
        eRequestedErrorSource := CAM_SOURCE_SLAVE_AXIS;
        udiRequestedMotionErrorID := fbSetPositionCutter.ErrorID;
    ELSIF fbMoveConveyor.Error
       OR (fbMoveConveyor.CommandAborted
           AND ((eState = CAM_STATE_STARTING_MASTER)
                OR (eState = CAM_STATE_CAMMING_IN)
                OR (eState = CAM_STATE_RUNNING))) THEN
        bRequestFault := TRUE;
        eRequestedApplicationError := CAM_ERROR_MASTER_MOVE;
        eRequestedErrorSource := CAM_SOURCE_MASTER_AXIS;
        udiRequestedMotionErrorID := fbMoveConveyor.ErrorID;
    ELSIF fbStopConveyor.Error THEN
        bRequestFault := TRUE;
        eRequestedApplicationError := CAM_ERROR_MASTER_STOP;
        eRequestedErrorSource := CAM_SOURCE_MASTER_AXIS;
        udiRequestedMotionErrorID := fbStopConveyor.ErrorID;
    ELSIF fbReturnCutter.Error OR fbReturnCutter.CommandAborted THEN
        bRequestFault := TRUE;
        eRequestedApplicationError := CAM_ERROR_SLAVE_RETURN;
        eRequestedErrorSource := CAM_SOURCE_SLAVE_AXIS;
        udiRequestedMotionErrorID := fbReturnCutter.ErrorID;
    ELSIF fbElectronicCam.bError THEN
        bRequestFault := TRUE;
        eRequestedApplicationError := fbElectronicCam.eApplicationError;
        eRequestedErrorSource := fbElectronicCam.eErrorSource;
        udiRequestedMotionErrorID := fbElectronicCam.udiErrorID;
    END_IF;
END_IF;

IF bRequestFault THEN
    IF NOT bFaultLatched THEN
        bFaultLatched := TRUE;
        eLatchedApplicationError := eRequestedApplicationError;
        eLatchedErrorSource := eRequestedErrorSource;
        udiLatchedMotionErrorID := udiRequestedMotionErrorID;
    END_IF;

    CASE eState OF
        CAM_STATE_STARTING_MASTER,
        CAM_STATE_CAMMING_IN,
        CAM_STATE_RUNNING:
            // Any runtime fault is stopped before entering the latched fault state.
            bMoveConveyorExecute := FALSE;
            bStopRequested := TRUE;
            bFaultStop := TRUE;
            eState := CAM_STATE_STOPPING_MASTER;
        CAM_STATE_STOPPING_MASTER:
            bFaultStop := TRUE;
        CAM_STATE_RELEASING_STOP,
        CAM_STATE_CAMMING_OUT,
        CAM_STATE_RETURNING_SLAVE,
        CAM_STATE_RESETTING:
            // Master is already stopped; finish the controlled recovery step.
    ELSE
        eState := CAM_STATE_FAULT;
    END_CASE;
END_IF;

// Scope signals are kept flat and use the NC cyclic set/actual values directly.
stScope.lrMasterSetPosition := AxisConveyor.NcToPlc.SetPos;
stScope.lrMasterActualPosition := AxisConveyor.NcToPlc.ActPos;
stScope.lrMasterSetVelocity := AxisConveyor.NcToPlc.SetVelo;
stScope.lrMasterActualVelocity := AxisConveyor.NcToPlc.ActVelo;
stScope.lrSlaveSetPosition := AxisCutter.NcToPlc.SetPos;
stScope.lrSlaveActualPosition := AxisCutter.NcToPlc.ActPos;
stScope.lrSlaveSetVelocity := AxisCutter.NcToPlc.SetVelo;
stScope.lrSlaveActualVelocity := AxisCutter.NcToPlc.ActVelo;

IF fbElectronicCam.bCamActive AND (stActiveRecipe.lrObjectPitch > 0.0) THEN
    stScope.lrMasterPhase := lrMasterPhase;
    lrSlaveCamPosition := AxisCutter.NcToPlc.SetPos - lrSlaveCycleOrigin;
    stScope.lrObjectRelativePosition :=
        lrSlaveCamPosition - stScope.lrMasterPhase;
ELSE
    stScope.lrMasterPhase := 0.0;
    stScope.lrObjectRelativePosition := 0.0;
END_IF;

IF eState = CAM_STATE_DISABLED THEN
    eProcessPhase := CAM_PHASE_DISABLED;
ELSIF stScope.lrMasterPhase < stActiveRecipe.lrBlendMasterDistance THEN
    eProcessPhase := CAM_PHASE_PREPARE;
ELSIF stScope.lrMasterPhase < stActiveRecipe.lrFirstEdgeStart THEN
    eProcessPhase := CAM_PHASE_APPROACH;
ELSIF stScope.lrMasterPhase < stDerived.lrFirstEdgeEnd THEN
    eProcessPhase := CAM_PHASE_FIRST_EDGE;
ELSIF stScope.lrMasterPhase < stDerived.lrExitBlendEnd THEN
    eProcessPhase := CAM_PHASE_EXIT_FIRST_EDGE;
ELSIF stScope.lrMasterPhase < stDerived.lrEntryBlendStart THEN
    eProcessPhase := CAM_PHASE_SYNCHRONOUS;
ELSIF stScope.lrMasterPhase < stActiveRecipe.lrSecondEdgeStart THEN
    eProcessPhase := CAM_PHASE_ENTER_SECOND_EDGE;
ELSIF stScope.lrMasterPhase < stDerived.lrSecondEdgeEnd THEN
    eProcessPhase := CAM_PHASE_SECOND_EDGE;
ELSIF stScope.lrMasterPhase < stActiveRecipe.lrReturnEndPhase THEN
    eProcessPhase := CAM_PHASE_RETURN;
ELSE
    eProcessPhase := CAM_PHASE_DWELL;
END_IF;

CASE eProcessPhase OF
    CAM_PHASE_FIRST_EDGE:
        stScope.lrExpectedSlaveVelocity :=
            stActiveRecipe.lrConveyorVelocity + stActiveRecipe.lrCutVelocity;
    CAM_PHASE_SYNCHRONOUS:
        stScope.lrExpectedSlaveVelocity := stActiveRecipe.lrConveyorVelocity;
    CAM_PHASE_SECOND_EDGE:
        stScope.lrExpectedSlaveVelocity :=
            stActiveRecipe.lrConveyorVelocity - stActiveRecipe.lrCutVelocity;
    CAM_PHASE_APPROACH,
    CAM_PHASE_EXIT_FIRST_EDGE,
    CAM_PHASE_ENTER_SECOND_EDGE,
    CAM_PHASE_RETURN:
        stScope.lrExpectedSlaveVelocity := AxisCutter.NcToPlc.SetVelo;
ELSE
    stScope.lrExpectedSlaveVelocity := 0.0;
END_CASE;

stStatus.eState := eState;
stStatus.eProcessPhase := eProcessPhase;
stStatus.bPowerEnabled := fbPowerConveyor.Status AND fbPowerCutter.Status;
stStatus.bReferenced := bReferenced;
stStatus.bRecipeLoaded := bRecipeLoaded;
stStatus.bCamActive := fbElectronicCam.bCamActive;
stStatus.bRunning := eState = CAM_STATE_RUNNING;
stStatus.bBusy := (eState <> CAM_STATE_DISABLED)
    AND (eState <> CAM_STATE_IDLE)
    AND (eState <> CAM_STATE_READY)
    AND (eState <> CAM_STATE_FAULT);
stStatus.eApplicationError := eLatchedApplicationError;
stStatus.eErrorSource := eLatchedErrorSource;
stStatus.udiMotionErrorID := udiLatchedMotionErrorID;
stStatus.lrCalculatedMaxSlaveVelocity := lrCalculatedMaxSlaveVelocity;
stStatus.lrCalculatedMaxSlaveAcceleration := lrCalculatedMaxSlaveAcceleration;
stStatus.lrCalculatedMaxSlaveJerk := lrCalculatedMaxSlaveJerk;
stStatus.lrCalculatedFaultStopSlaveAcceleration :=
    lrCalculatedFaultStopSlaveAcceleration;
stStatus.lrCalculatedFaultStopSlaveJerk :=
    lrCalculatedFaultStopSlaveJerk;

stScope.eMachineState := eState;
stScope.eProcessPhase := eProcessPhase;
stScope.bCamActive := fbElectronicCam.bCamActive;
stScope.bRecipeLoaded := bRecipeLoaded;
stScope.eApplicationError := eLatchedApplicationError;
stScope.udiMotionErrorID := udiLatchedMotionErrorID;

END_FUNCTION_BLOCK

// ---- POUs/Cam/FB_CamRecipeValidator.TcPOU
FUNCTION_BLOCK FB_CamRecipeValidator
VAR_INPUT
    bExecute : BOOL;
    stRecipe : ST_CamRecipe;
END_VAR
VAR_OUTPUT
    bDone : BOOL;
    bValid : BOOL;
    bError : BOOL;
    eError : E_CamApplicationError;
    stDerived : ST_CamDerivedGeometry;
END_VAR
VAR
    rtExecute : R_TRIG;
END_VAR
VAR CONSTANT
    c_lrPlcCycleSeconds : LREAL := 0.01;
    c_lrSaneUpperBound : LREAL := 1.0E9;
END_VAR

rtExecute(CLK := bExecute);
bDone := FALSE;

IF rtExecute.Q THEN
    bValid := FALSE;
    bError := FALSE;
    eError := CAM_ERROR_NONE;

    // The paired comparisons also reject NaN and infinity-like values.
    IF NOT ((stRecipe.lrObjectPitch > 0.0)
       AND (stRecipe.lrObjectPitch < c_lrSaneUpperBound)) THEN
        eError := CAM_ERROR_RECIPE_PITCH;
    ELSIF NOT ((stRecipe.lrConveyorVelocity > 0.0)
       AND (stRecipe.lrConveyorVelocity < c_lrSaneUpperBound)) THEN
        eError := CAM_ERROR_RECIPE_CONVEYOR_VELOCITY;
    ELSIF NOT ((stRecipe.lrCutVelocity > 0.0)
       AND (stRecipe.lrCutVelocity < stRecipe.lrConveyorVelocity)) THEN
        eError := CAM_ERROR_RECIPE_CUT_VELOCITY;
    ELSIF NOT ((stRecipe.lrObjectEdgeLength > 0.0)
       AND (stRecipe.lrObjectEdgeLength < c_lrSaneUpperBound)
       AND (stRecipe.lrBlendMasterDistance > 0.0)
       AND (stRecipe.lrBlendMasterDistance < c_lrSaneUpperBound)
       AND (stRecipe.lrFirstEdgeStart > 0.0)
       AND (stRecipe.lrFirstEdgeStart < c_lrSaneUpperBound)
       AND (stRecipe.lrSecondEdgeStart > 0.0)
       AND (stRecipe.lrSecondEdgeStart < c_lrSaneUpperBound)
       AND (stRecipe.lrReturnEndPhase > 0.0)
       AND (stRecipe.lrReturnEndPhase < c_lrSaneUpperBound)) THEN
        eError := CAM_ERROR_RECIPE_EDGE_LENGTH;
    ELSIF NOT ((stRecipe.lrMasterAcceleration > 0.0)
       AND (stRecipe.lrMasterAcceleration < c_lrSaneUpperBound)
       AND (stRecipe.lrMasterDeceleration > 0.0)
       AND (stRecipe.lrMasterDeceleration < c_lrSaneUpperBound)
       AND (stRecipe.lrMasterJerk > 0.0)
       AND (stRecipe.lrMasterJerk < c_lrSaneUpperBound)
       AND (stRecipe.lrRecoveryVelocity > 0.0)
       AND (stRecipe.lrRecoveryVelocity < c_lrSaneUpperBound)
       AND (stRecipe.lrRecoveryAcceleration > 0.0)
       AND (stRecipe.lrRecoveryAcceleration < c_lrSaneUpperBound)
       AND (stRecipe.lrRecoveryDeceleration > 0.0)
       AND (stRecipe.lrRecoveryDeceleration < c_lrSaneUpperBound)
       AND (stRecipe.lrRecoveryJerk > 0.0)
       AND (stRecipe.lrRecoveryJerk < c_lrSaneUpperBound)
       AND (stRecipe.lrPositionTolerance > 0.0)
       AND (stRecipe.lrPositionTolerance < c_lrSaneUpperBound)
       AND (stRecipe.lrMaxSlaveVelocity > 0.0)
       AND (stRecipe.lrMaxSlaveVelocity < c_lrSaneUpperBound)
       AND (stRecipe.lrMaxSlaveAcceleration > 0.0)
       AND (stRecipe.lrMaxSlaveAcceleration < c_lrSaneUpperBound)
       AND (stRecipe.lrMaxSlaveJerk > 0.0)
       AND (stRecipe.lrMaxSlaveJerk < c_lrSaneUpperBound)) THEN
        eError := CAM_ERROR_RECIPE_DYNAMICS;
    ELSE
        stDerived.lrCutMasterDistance :=
            stRecipe.lrObjectEdgeLength * stRecipe.lrConveyorVelocity
            / stRecipe.lrCutVelocity;
        stDerived.lrFirstSlope :=
            1.0 + stRecipe.lrCutVelocity / stRecipe.lrConveyorVelocity;
        stDerived.lrSecondSlope :=
            1.0 - stRecipe.lrCutVelocity / stRecipe.lrConveyorVelocity;
        stDerived.lrFirstEdgeEnd :=
            stRecipe.lrFirstEdgeStart + stDerived.lrCutMasterDistance;
        stDerived.lrExitBlendEnd :=
            stDerived.lrFirstEdgeEnd + stRecipe.lrBlendMasterDistance;
        stDerived.lrEntryBlendStart :=
            stRecipe.lrSecondEdgeStart - stRecipe.lrBlendMasterDistance;
        stDerived.lrSecondEdgeEnd :=
            stRecipe.lrSecondEdgeStart + stDerived.lrCutMasterDistance;
        stDerived.lrFirstStartY := stRecipe.lrFirstEdgeStart;
        stDerived.lrFirstEndY := stDerived.lrFirstStartY
            + stDerived.lrFirstSlope * stDerived.lrCutMasterDistance;
        stDerived.lrExitEndY := stDerived.lrFirstEndY
            + 0.5 * (stDerived.lrFirstSlope + 1.0)
            * stRecipe.lrBlendMasterDistance;
        stDerived.lrClearanceRelative :=
            stDerived.lrExitEndY - stDerived.lrExitBlendEnd;
        stDerived.lrEntryStartY :=
            stDerived.lrEntryBlendStart + stDerived.lrClearanceRelative;
        stDerived.lrSecondStartY :=
            stRecipe.lrSecondEdgeStart + stRecipe.lrObjectEdgeLength;
        stDerived.lrSecondEndY := stDerived.lrSecondStartY
            + stDerived.lrSecondSlope * stDerived.lrCutMasterDistance;

        // Symmetric jerk-limited stop distance from steady conveyor speed.
        IF stRecipe.lrConveyorVelocity >=
           (stRecipe.lrMasterDeceleration * stRecipe.lrMasterDeceleration
            / stRecipe.lrMasterJerk) THEN
            stDerived.lrMasterStopDistance :=
                0.5 * stRecipe.lrConveyorVelocity
                * (stRecipe.lrConveyorVelocity / stRecipe.lrMasterDeceleration
                   + stRecipe.lrMasterDeceleration / stRecipe.lrMasterJerk);
        ELSE
            stDerived.lrMasterStopDistance :=
                stRecipe.lrConveyorVelocity
                * SQRT(stRecipe.lrConveyorVelocity / stRecipe.lrMasterJerk);
        END_IF;
        stDerived.lrStopWindowMargin :=
            2.0 * c_lrPlcCycleSeconds * stRecipe.lrConveyorVelocity;

        IF stRecipe.lrFirstEdgeStart <= stRecipe.lrBlendMasterDistance THEN
            eError := CAM_ERROR_RECIPE_PHASE_ORDER;
        ELSIF stDerived.lrExitBlendEnd >= stDerived.lrEntryBlendStart THEN
            eError := CAM_ERROR_RECIPE_SYNC_SPACE;
        ELSIF (stDerived.lrSecondEdgeEnd >= stRecipe.lrReturnEndPhase)
           OR (stRecipe.lrReturnEndPhase >= stRecipe.lrObjectPitch) THEN
            eError := CAM_ERROR_RECIPE_RETURN_SPACE;
        ELSIF (stDerived.lrMasterStopDistance
               + stDerived.lrStopWindowMargin)
              > (stRecipe.lrObjectPitch - stRecipe.lrReturnEndPhase) THEN
            eError := CAM_ERROR_RECIPE_DYNAMICS;
        ELSE
            bValid := TRUE;
        END_IF;
    END_IF;

    bError := NOT bValid;
    bDone := TRUE;
END_IF;

END_FUNCTION_BLOCK

// ---- POUs/Cam/FB_CamProfileBuilder.TcPOU
FUNCTION_BLOCK FB_CamProfileBuilder
VAR_INPUT
    bExecute : BOOL;
    stRecipe : ST_CamRecipe;
    stDerived : ST_CamDerivedGeometry;
END_VAR
VAR_OUTPUT
    bDone : BOOL;
    aPoints : ARRAY[1..10] OF MC_MotionFunctionPoint;
    stCamRef : MC_CAM_REF;
END_VAR
VAR
    rtExecute : R_TRIG;
END_VAR

rtExecute(CLK := bExecute);
bDone := FALSE;

IF rtExecute.Q THEN
    aPoints[1] := F_MakeCamPoint(1, MOTIONFUNCTYPE_POLYNOM1,
        MOTIONPOINTTYPE_REST, 1, 0.0, 0.0, 0.0);
    aPoints[2] := F_MakeCamPoint(2, MOTIONFUNCTYPE_POLYNOM5_MM,
        MOTIONPOINTTYPE_REST, 1,
        stRecipe.lrBlendMasterDistance, 0.0, 0.0);
    aPoints[3] := F_MakeCamPoint(3, MOTIONFUNCTYPE_POLYNOM1,
        MOTIONPOINTTYPE_VELOCITY, 1, stRecipe.lrFirstEdgeStart,
        stDerived.lrFirstStartY, stDerived.lrFirstSlope);
    aPoints[4] := F_MakeCamPoint(4, MOTIONFUNCTYPE_POLYNOM5_MM,
        MOTIONPOINTTYPE_VELOCITY, 1, stDerived.lrFirstEdgeEnd,
        stDerived.lrFirstEndY, stDerived.lrFirstSlope);
    aPoints[5] := F_MakeCamPoint(5, MOTIONFUNCTYPE_POLYNOM1,
        MOTIONPOINTTYPE_VELOCITY, 1, stDerived.lrExitBlendEnd,
        stDerived.lrExitEndY, 1.0);
    aPoints[6] := F_MakeCamPoint(6, MOTIONFUNCTYPE_POLYNOM5_MM,
        MOTIONPOINTTYPE_VELOCITY, 1, stDerived.lrEntryBlendStart,
        stDerived.lrEntryStartY, 1.0);
    aPoints[7] := F_MakeCamPoint(7, MOTIONFUNCTYPE_POLYNOM1,
        MOTIONPOINTTYPE_VELOCITY, 1, stRecipe.lrSecondEdgeStart,
        stDerived.lrSecondStartY, stDerived.lrSecondSlope);
    aPoints[8] := F_MakeCamPoint(8, MOTIONFUNCTYPE_POLYNOM5_MM,
        MOTIONPOINTTYPE_VELOCITY, 1, stDerived.lrSecondEdgeEnd,
        stDerived.lrSecondEndY, stDerived.lrSecondSlope);
    aPoints[9] := F_MakeCamPoint(9, MOTIONFUNCTYPE_POLYNOM1,
        MOTIONPOINTTYPE_REST, 1, stRecipe.lrReturnEndPhase, 0.0, 0.0);
    aPoints[10] := F_MakeCamPoint(10, MOTIONFUNCTYPE_NOTDEF,
        MOTIONPOINTTYPE_REST, 0, stRecipe.lrObjectPitch, 0.0, 0.0);

    stCamRef.pArray := ADR(aPoints);
    stCamRef.ArraySize := SIZEOF(aPoints);
    stCamRef.TableType := MC_TABLETYPE_MOTIONFUNCTION;
    stCamRef.NoOfRows := 10;
    stCamRef.NoOfColumns := 1;
    bDone := TRUE;
END_IF;

END_FUNCTION_BLOCK

// ---- POUs/Cam/F_MakeCamPoint.TcPOU
FUNCTION F_MakeCamPoint : MC_MotionFunctionPoint
VAR_INPUT
    udiPointIndex : UDINT;
    eFunctionType : MC_MotionFunctionType;
    ePointType : MC_MotionPointType;
    udiRelIndexNextPoint : UDINT;
    lrMasterPos : LREAL;
    lrSlavePos : LREAL;
    lrSlaveVelo : LREAL;
END_VAR

F_MakeCamPoint.PointIndex := udiPointIndex;
F_MakeCamPoint.FunctionType := eFunctionType;
F_MakeCamPoint.PointType := ePointType;
F_MakeCamPoint.RelIndexNextPoint := udiRelIndexNextPoint;
F_MakeCamPoint.MasterPos := lrMasterPos;
F_MakeCamPoint.SlavePos := lrSlavePos;
F_MakeCamPoint.SlaveVelo := lrSlaveVelo;
F_MakeCamPoint.SlaveAcc := 0.0;
F_MakeCamPoint.SlaveJerk := 0.0;

END_FUNCTION

// ---- POUs/Cam/FB_ElectronicCam.TcPOU
FUNCTION_BLOCK FB_ElectronicCam
VAR_INPUT
    bLoad : BOOL;
    bCouple : BOOL;
    bDecouple : BOOL;
    bReset : BOOL;
    nCamTableId : MC_CAM_ID := 1;
END_VAR
VAR_IN_OUT
    Master : AXIS_REF;
    Slave : AXIS_REF;
    CamTable : MC_CAM_REF;
END_VAR
VAR_OUTPUT
    bLoadDone : BOOL;
    bCoupleDone : BOOL;
    bDecoupleDone : BOOL;
    bBusy : BOOL;
    bCamActive : BOOL;
    bError : BOOL;
    eApplicationError : E_CamApplicationError;
    eErrorSource : E_CamErrorSource;
    udiErrorID : UDINT;
    stCharacteristics : MC_TableCharacValues;
END_VAR
VAR
    rtLoad : R_TRIG;
    rtCouple : R_TRIG;
    rtDecouple : R_TRIG;
    fbTableSelect : MC_CamTableSelect;
    fbCharacteristics : MC_ReadCamTableCharacteristics;
    fbCamIn : MC_CamIn;
    fbCamOut : MC_CamOut;
    stCamInOptions : ST_CamInOptions;
    stCharacteristicsOptions : ST_ReadCamTableCharacteristicsOptions;
    stCamOutOptions : ST_CamOutOptions;
    bTableSelectExecute : BOOL;
    bCharacteristicsExecute : BOOL;
    bCamInExecute : BOOL;
    bCamOutExecute : BOOL;
    usiLoadState : USINT;
END_VAR

rtLoad(CLK := bLoad);
rtCouple(CLK := bCouple);
rtDecouple(CLK := bDecouple);

bLoadDone := FALSE;
bCoupleDone := FALSE;
bDecoupleDone := FALSE;

IF bReset THEN
    bTableSelectExecute := FALSE;
    bCharacteristicsExecute := FALSE;
    bCamInExecute := FALSE;
    bCamOutExecute := FALSE;
    usiLoadState := 0;
    bError := FALSE;
    eApplicationError := CAM_ERROR_NONE;
    eErrorSource := CAM_SOURCE_NONE;
    udiErrorID := 0;
END_IF;

// Accept at most one command when the wrapper is idle.
IF NOT bReset AND NOT bError THEN
    IF rtLoad.Q
       AND (usiLoadState = 0)
       AND NOT bCamInExecute
       AND NOT bCamOutExecute
       AND NOT bCamActive THEN
        usiLoadState := 10;
        bTableSelectExecute := TRUE;
    ELSIF rtCouple.Q
       AND (usiLoadState = 0)
       AND NOT bCamInExecute
       AND NOT bCamOutExecute
       AND NOT bCamActive THEN
        bCamInExecute := TRUE;
    ELSIF rtDecouple.Q
       AND (usiLoadState = 0)
       AND NOT bCamInExecute
       AND NOT bCamOutExecute
       AND bCamActive THEN
        bCamOutExecute := TRUE;
    END_IF;
END_IF;

fbTableSelect(
    Execute := bTableSelectExecute,
    Periodic := TRUE,
    MasterAbsolute := FALSE,
    SlaveAbsolute := FALSE,
    CamTableID := nCamTableId,
    Master := Master,
    Slave := Slave,
    CamTable := CamTable);
fbCharacteristics(
    Execute := bCharacteristicsExecute,
    CamTableID := nCamTableId,
    Options := stCharacteristicsOptions,
    CamTableCharac := stCharacteristics);
fbCamIn(
    Execute := bCamInExecute,
    MasterOffset := 0.0,
    SlaveOffset := 0.0,
    MasterScaling := 1.0,
    SlaveScaling := 1.0,
    StartMode := MC_STARTMODE_RELATIVE,
    CamTableID := nCamTableId,
    BufferMode := MC_Aborting,
    Options := stCamInOptions,
    Master := Master,
    Slave := Slave);
fbCamOut(
    Execute := bCamOutExecute,
    Options := stCamOutOptions,
    Slave := Slave);

IF NOT bReset THEN
    // Preserve the first NC error until the caller resets this wrapper.
    IF NOT bError THEN
        IF fbTableSelect.Error THEN
            bError := TRUE;
            eApplicationError := CAM_ERROR_CAM_LOAD;
            eErrorSource := CAM_SOURCE_TABLE_LOAD;
            udiErrorID := fbTableSelect.ErrorID;
        ELSIF fbCharacteristics.Error THEN
            bError := TRUE;
            eApplicationError := CAM_ERROR_CAM_CHARACTERISTICS;
            eErrorSource := CAM_SOURCE_TABLE_CHARACTERISTICS;
            udiErrorID := fbCharacteristics.ErrorID;
        ELSIF fbCamIn.Error OR fbCamIn.CommandAborted THEN
            bError := TRUE;
            eApplicationError := CAM_ERROR_CAM_IN;
            eErrorSource := CAM_SOURCE_CAM_IN;
            udiErrorID := fbCamIn.ErrorID;
        ELSIF fbCamOut.Error THEN
            bError := TRUE;
            eApplicationError := CAM_ERROR_CAM_OUT;
            eErrorSource := CAM_SOURCE_CAM_OUT;
            udiErrorID := fbCamOut.ErrorID;
        END_IF;
    END_IF;

    IF bError THEN
        bTableSelectExecute := FALSE;
        bCharacteristicsExecute := FALSE;
        bCamInExecute := FALSE;
        bCamOutExecute := FALSE;
        usiLoadState := 0;
    ELSE
        CASE usiLoadState OF
            10:
                IF fbTableSelect.Done THEN
                    bTableSelectExecute := FALSE;
                    bCharacteristicsExecute := TRUE;
                    usiLoadState := 20;
                END_IF;

            20:
                IF fbCharacteristics.Done THEN
                    bCharacteristicsExecute := FALSE;
                    usiLoadState := 0;
                    bLoadDone := TRUE;
                END_IF;
        END_CASE;

        IF fbCamIn.InSync THEN
            bCamInExecute := FALSE;
            bCamActive := TRUE;
            bCoupleDone := TRUE;
        END_IF;

        IF fbCamOut.Done THEN
            bCamOutExecute := FALSE;
            bCamActive := FALSE;
            bDecoupleDone := TRUE;
        END_IF;
    END_IF;
END_IF;

bBusy := (usiLoadState <> 0)
    OR bTableSelectExecute
    OR bCharacteristicsExecute
    OR bCamInExecute
    OR bCamOutExecute
    OR fbTableSelect.Busy
    OR fbCharacteristics.Busy
    OR fbCamIn.Busy
    OR fbCamOut.Busy;

END_FUNCTION_BLOCK

// ---- POUs/Axis_test/Axis_test.TcPOU
PROGRAM Axis_test
VAR
    // Online commands: bMoveAbsolute and bStop are rising-edge commands.
    bPower : BOOL := FALSE;
    bMoveAbsolute : BOOL := FALSE;
    bStop : BOOL := FALSE;
	bReset : BOOL := FALSE;

    // Values use the engineering unit configured for the selected NC axis.
    lrTargetPosition : LREAL := 0.0;
    lrVelocity : LREAL := 5.0;
    lrAcceleration : LREAL := 20.0;
    lrDeceleration : LREAL := 20.0;
    lrJerk : LREAL := 100.0;

    // Online diagnostics.
    bPowerStatus : BOOL;
    bMoveBusy : BOOL;
    bMoveDone : BOOL;
    bStopDone : BOOL;
    bError : BOOL;
    udiErrorID : UDINT;
    lrActualPosition : LREAL;

    fbAxisTest : FB_AxisPositionTest;
END_VAR

fbAxisTest(
    bPower := bPower,
    bMoveAbsolute := bMoveAbsolute,
	bReset := bReset,
    bStop := bStop,
    lrTargetPosition := lrTargetPosition,
    lrVelocity := lrVelocity,
    lrAcceleration := lrAcceleration,
    lrDeceleration := lrDeceleration,
    lrJerk := lrJerk,
    // Change only this line to select another test axis.
    Axis := GVL_Motion.gAxisConveyor,
    bPowerStatus => bPowerStatus,
    bMoveBusy => bMoveBusy,
    bMoveDone => bMoveDone,
    bStopDone => bStopDone,
    bError => bError,
    udiErrorID => udiErrorID,
    lrActualPosition => lrActualPosition);

END_PROGRAM

// ---- POUs/Axis_test/FB_AxisPositionTest.TcPOU
FUNCTION_BLOCK FB_AxisPositionTest
VAR_INPUT
    bPower : BOOL;
    bMoveAbsolute : BOOL;
	bReset: BOOL;
    bStop : BOOL;
    lrTargetPosition : LREAL;
    lrVelocity : LREAL;
    lrAcceleration : LREAL;
    lrDeceleration : LREAL;
    lrJerk : LREAL;
END_VAR
VAR_IN_OUT
    Axis : AXIS_REF;
END_VAR
VAR_OUTPUT
    bPowerStatus : BOOL;
    bMoveBusy : BOOL;
    bMoveDone : BOOL;
    bStopDone : BOOL;
    bError : BOOL;
    udiErrorID : UDINT;
    lrActualPosition : LREAL;
END_VAR
VAR
    fbPower : MC_Power;
	fbReset : MC_Reset;
    fbMoveAbsolute : MC_MoveAbsolute;
    fbStop : MC_Stop;
    stPowerOptions : ST_PowerOptions;
    stMoveOptions : ST_MoveOptions;
    stStopOptions : ST_MoveOptions;
END_VAR

Axis.ReadStatus();

fbPower(
    Enable := bPower,
    Enable_Positive := TRUE,
    Enable_Negative := TRUE,
    Override := 100.0,
    BufferMode := MC_Aborting,
    Options := stPowerOptions,
    Axis := Axis);

fbMoveAbsolute(
    Execute := bMoveAbsolute AND NOT bStop,
    Position := lrTargetPosition,
    Velocity := lrVelocity,
    Acceleration := lrAcceleration,
    Deceleration := lrDeceleration,
    Jerk := lrJerk,
    BufferMode := MC_Aborting,
    Options := stMoveOptions,
    Axis := Axis);

fbReset(Axis := Axis,Execute := bReset);

fbStop(
    Execute := bStop,
    Deceleration := lrDeceleration,
    Jerk := lrJerk,
    Options := stStopOptions,
    Axis := Axis);

bPowerStatus := fbPower.Status;
bMoveBusy := fbMoveAbsolute.Busy;
bMoveDone := fbMoveAbsolute.Done;
bStopDone := fbStop.Done;
bError := fbPower.Error OR fbMoveAbsolute.Error OR fbStop.Error;
IF fbPower.Error THEN
    udiErrorID := fbPower.ErrorID;
ELSIF fbMoveAbsolute.Error THEN
    udiErrorID := fbMoveAbsolute.ErrorID;
ELSIF fbStop.Error THEN
    udiErrorID := fbStop.ErrorID;
ELSE
    udiErrorID := 0;
END_IF;
lrActualPosition := Axis.NcToPlc.ActPos;

END_FUNCTION_BLOCK

// ---- POUs/MAIN.TcPOU
PROGRAM MAIN
VAR
    fbCamMachine : FB_CamMachine;
END_VAR

fbCamMachine(
    stCommands := GVL_CamControl.stCommands,
    stRecipe := GVL_CamControl.stRecipe,
    AxisConveyor := GVL_Motion.gAxisConveyor,
    AxisCutter := GVL_Motion.gAxisCutter,
    stStatus => GVL_CamControl.stStatus,
    stScope => GVL_CamControl.stScope);

END_PROGRAM
